# EPICS substitutions: examples/PSI/plugins/cpp_logic/examples/cpp_logic_minimal_el1252/cfg/libmain.so_cpp_logic.subs
# Auto-generated C++ logic substitutions
# Logic: cpp_logic_minimal_uint64
global { P = "$(P)" PORT = "$(PORT)" }

file ecmcCppLogicAi.template {
  pattern { REC,                    ASYN_OPT,                                 PARAM,                           DESC,                            DTYP,        SCAN       }
  { "main-timestampLatchPositive01","/TYPE=asynFloat64/CMD=UINT64TOFLOAT64/", "main.timestampLatchPositive01", "main.timestampLatchPositive01", asynFloat64, "I/O Intr" }
}
